// SIMATIC S7-200 project (STEP 7-Micro/WIN), CPU 224 CN REL 02.01

SYMBOL_TABLE USUARIO1
SB_2             I1.2     // Pulsador de paro
SB_1             I1.3     // Pulsador de marcha
QS               I1.4     // Zeta de emergencia
SA               I1.5     // Selector de modo
HL1              Q0.7     // Piloto amarillo
HL2              Q1.0     // Piloto verde
HL3              Q1.1     // Piloto rojo
END_SYMBOL_TABLE

ORGANIZATION_BLOCK PRINCIPAL:OB1
TITLE=COMENTARIOS DEL PROGRAMA
BEGIN
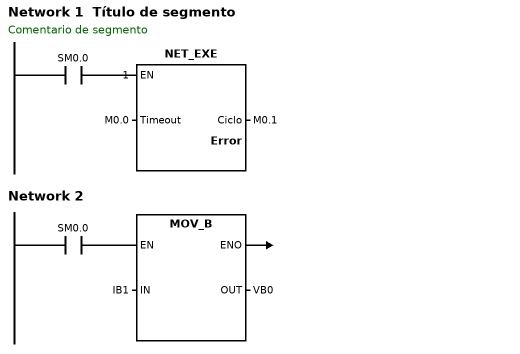
Network 1 // Título de segmento
// Comentario de segmento
// (network saved uncompiled; LAD cells follow)
// row 0: c0 -| |- SM0.0  c1 [NET_EXE Error EN:=1, Timeout:=M0.0, Ciclo=>M0.1]
// row 1: c1 [box]
Network 2
// (network saved uncompiled; LAD cells follow)
// row 0: c0 -| |- SM0.0  c1 [MOV_B EN:=power@row0, IN:=IB1, ENO=>power, OUT=>VB0]  c2 ->
// row 1: c1 [box]
END_ORGANIZATION_BLOCK

// SBR1: protected block, not included
